(*
    Pneumatic actuator, single or double acting, ported from the legacy
    FB_MotionPneumaticActuator. Implements I_PneumaticActuator. The limit switch state, the
    insert and retract exclusion and the output timeout come from FB_PneumaticCore, which
    FB_MPA uses as well.

    Position state from the limit switches (in = inserted LS, out = retracted LS):
        in AND out         INVALID
        NOT in AND out     RETRACTED
        in AND NOT out     INSERTED
        NOT in AND NOT out MOVING
    bDone: the commanded direction has reached its limit switch. bBusy: a command
    is active and its limit switch is not reached. xMPS_OK is TRUE only when the
    state is RETRACTED or INSERTED. The fast fault (device 'MPA', type code
    E_MotionFFType.PNEUMATIC_MOVE) trips when xMPS_OK is FALSE.

    Insert and retract requests are mutually exclusive: both set at once clears both.
    Single acting: ibSingleCntrl TRUE and ibCntrlHold TRUE keeps the output on after
    arrival. Double acting: both FALSE, the output drops once the limit switch of the
    commanded direction has been active for LimitSwitchLatchDuration (default 1 s).
    An output that does not reach its limit switch within TimeoutDuration (default
    10 s) sets bError and sErrorMessage until bReset is set.

    Legacy behaviour kept as is: ibPMPS_OK and ibOverrideInterlock are unused (PMPS
    permission is not implemented), and LogEvents (legacy ACT_Logger) is never called by the body.
*)
FUNCTION_BLOCK FB_PneumaticActuator IMPLEMENTS I_PneumaticActuator
VAR_INPUT
    // Actuator can be inserted
    ibInsertOK : BOOL;
    // Actuator can be retracted
    ibRetractOK : BOOL;
    // To be linked to the arbiter bit (unused, as in the legacy FB)
    ibPMPS_OK : BOOL;
    // TRUE if the actuator needs one output (single acting), FALSE if it needs two
    ibSingleCntrl : BOOL;
    // Output must keep its value. TRUE for single acting, FALSE for double acting
    ibCntrlHold : BOOL;
    // If TRUE interlocks are ignored (unused, as in the legacy FB)
    ibOverrideInterlock : BOOL;
    {attribute 'pytmc' := '
    pv: FFO_Reset
    '}
    i_xReset : BOOL;
    {attribute 'pytmc' := '
    pv: FFO_AutoReset
    '}
    i_xAutoReset : BOOL;
END_VAR
VAR_OUTPUT
    {attribute 'pytmc' := '
    pv:
    '}
    stPneumaticActuator : ST_PneumaticActuator;
    {attribute 'pytmc' := '
     pv: MPS_OK
     field: ZNAM FALSE
     field: ONAM TRUE
     field: DESC TRUE if MPS signal is OK
    '}
    xMPS_OK : BOOL;
END_VAR
VAR
    // Fast fault output the fault is raised on
    fbFFHWO : REFERENCE TO FB_HardwareFFOutput;
    // Fault occurs while the actuator is not at a limit switch
    fbFF : FB_FastFault := (
        i_DevName := 'MPA',
        i_Desc := 'Fault occurs when the device is moving',
        i_TypeCode := E_MotionFFType.PNEUMATIC_MOVE);

    ftInit : R_TRIG;
    bFirstPass : BOOL;

    // Shared behaviour of the pneumatic actuator blocks
    fbCore : FB_PneumaticCore;
    // Time an output may stay on without reaching its limit switch
    tTimeOutDuration : TIME := T#10S;
    // Time a limit switch must stay active before a double acting output drops
    tLimitSwitchLatchDuration : TIME := T#1S;
    tonInsertLimitSwitch : TON;
    tonRetractLimitSwitch : TON;

    fbLogger : FB_LogMessage := (eSubsystem := E_SubSystem.MOTION);
    ePrevState : E_PnuematicActuatorPositionState;
    ftAction : R_TRIG;

    i_xInsertedLS AT %I* : BOOL;
    i_xRetractedLS AT %I* : BOOL;
    q_xInsert_DO AT %Q* : BOOL;
    q_xRetract_DO AT %Q* : BOOL;
END_VAR

IF NOT __ISVALIDREF(fbFFHWO) THEN
    RETURN;
END_IF

ftInit(CLK := TRUE, Q => bFirstPass);
IF bFirstPass THEN
    stPneumaticActuator.eState := E_PnuematicActuatorPositionState.INVALID;
    stPneumaticActuator.bRetractCmd := FALSE;
    stPneumaticActuator.bInsertCmd := FALSE;
END_IF

UpdateIO();

// Position state from the limit switches
// The output bits are those of the previous scan, so the timeout is reported one scan late
fbCore(
    bInLimitSwitch := stPneumaticActuator.bInLimitSwitch,
    bOutLimitSwitch := stPneumaticActuator.bOutLimitSwitch,
    bInsertOutput := stPneumaticActuator.bInsertOutput,
    bRetractOutput := stPneumaticActuator.bRetractOutput,
    tTimeout := tTimeOutDuration,
    eState => stPneumaticActuator.eState);

stPneumaticActuator.bDone := (stPneumaticActuator.bRetractCmd AND stPneumaticActuator.eState = E_PnuematicActuatorPositionState.RETRACTED)
    OR (stPneumaticActuator.bInsertCmd AND stPneumaticActuator.eState = E_PnuematicActuatorPositionState.INSERTED);
stPneumaticActuator.bBusy := (stPneumaticActuator.bRetractCmd AND stPneumaticActuator.eState <> E_PnuematicActuatorPositionState.RETRACTED)
    OR (stPneumaticActuator.bInsertCmd AND stPneumaticActuator.eState <> E_PnuematicActuatorPositionState.INSERTED);

// MPS faults when the actuator is in motion
xMPS_OK := (stPneumaticActuator.eState = E_PnuematicActuatorPositionState.RETRACTED)
    OR (stPneumaticActuator.eState = E_PnuematicActuatorPositionState.INSERTED);

// PMPS permission: yet to be implemented

// Insert and retract requests cannot both be active
IF stPneumaticActuator.bInsertCmd AND stPneumaticActuator.bRetractCmd THEN
    stPneumaticActuator.bInsertCmd := FALSE;
    stPneumaticActuator.bRetractCmd := FALSE;
END_IF

// Redundant: clear the opposite output and request when one output is active
IF stPneumaticActuator.bInsertOutput THEN
    stPneumaticActuator.bRetractOutput := FALSE;
    stPneumaticActuator.bRetractCmd := FALSE;
END_IF
IF stPneumaticActuator.bRetractOutput THEN
    stPneumaticActuator.bInsertOutput := FALSE;
    stPneumaticActuator.bInsertCmd := FALSE;
END_IF

stPneumaticActuator.bRetractOutput := stPneumaticActuator.bRetractOK
    AND stPneumaticActuator.bRetractCmd
    AND NOT stPneumaticActuator.bInsertCmd;
stPneumaticActuator.bInsertOutput := stPneumaticActuator.bInsertOK
    AND stPneumaticActuator.bInsertCmd
    AND NOT stPneumaticActuator.bRetractCmd;

// Double acting: drop the output once the actuator is seated in its limit switch
IF NOT ibSingleCntrl AND NOT ibCntrlHold THEN
    IF stPneumaticActuator.bRetractCmd
        AND stPneumaticActuator.bOutLimitSwitch
        AND tonRetractLimitSwitch.Q THEN
        stPneumaticActuator.bRetractOutput := FALSE;
    END_IF
    IF stPneumaticActuator.bInsertCmd
        AND stPneumaticActuator.bInLimitSwitch
        AND tonInsertLimitSwitch.Q THEN
        stPneumaticActuator.bInsertOutput := FALSE;
    END_IF
END_IF

tonInsertLimitSwitch(IN := stPneumaticActuator.bInLimitSwitch, PT := tLimitSwitchLatchDuration);
tonRetractLimitSwitch(IN := stPneumaticActuator.bOutLimitSwitch, PT := tLimitSwitchLatchDuration);

// Moving position timeout
IF fbCore.bInsertTimedOut THEN
    stPneumaticActuator.bError := TRUE;
    stPneumaticActuator.sErrorMessage := 'Actuator insert timeout';
ELSIF fbCore.bRetractTimedOut THEN
    stPneumaticActuator.bError := TRUE;
    stPneumaticActuator.sErrorMessage := 'Actuator retract timeout';
END_IF
stPneumaticActuator.bError R= stPneumaticActuator.bReset;

fbFF(
    i_xOK := xMPS_OK,
    i_xReset := i_xReset,
    i_xAutoReset := i_xAutoReset,
    io_fbFFHWO := fbFFHWO
);

UpdateIO();

PROPERTY Busy : BOOL
GET
Busy := stPneumaticActuator.bBusy;
END_GET
END_PROPERTY

(* Rebinds the fast fault output. Call from the CallAfterInit of an enclosing FB. *)
METHOD CallAfterInitActuator
VAR_INPUT
    fbFFHWO : REFERENCE TO FB_HardwareFFOutput;
END_VAR
THIS^.fbFFHWO REF= fbFFHWO;
END_METHOD

PROPERTY Done : BOOL
GET
Done := stPneumaticActuator.bDone;
END_GET
END_PROPERTY

PROPERTY Error : BOOL
GET
Error := stPneumaticActuator.bError;
END_GET
END_PROPERTY

// Text of the active timeout error
PROPERTY ErrorMessage : STRING
GET
ErrorMessage := stPneumaticActuator.sErrorMessage;
END_GET
END_PROPERTY

// Error reset request, the same bit as the reset PV
PROPERTY ErrorReset : BOOL
GET
ErrorReset := stPneumaticActuator.bReset;
END_GET
SET
stPneumaticActuator.bReset := ErrorReset;
END_SET
END_PROPERTY

(* Stores the mandatory fast fault output at instantiation. *)
METHOD FB_Init : BOOL
VAR_INPUT
    // TRUE: the retain variables are initialized (reset warm / reset cold)
    bInitRetains : BOOL;
    // TRUE: the instance will be copied to the copy code afterward (online change)
    bInCopyCode : BOOL;
    fbFFHWO : REFERENCE TO FB_HardwareFFOutput;
END_VAR
THIS^.fbFFHWO REF= fbFFHWO;
END_METHOD

METHOD Insert
VAR_INPUT
END_VAR
stPneumaticActuator.bInsertCmd := TRUE;
END_METHOD

// Insert request, the same bit Insert() raises. Write FALSE to clear it
PROPERTY InsertCmd : BOOL
GET
InsertCmd := stPneumaticActuator.bInsertCmd;
END_GET
SET
stPneumaticActuator.bInsertCmd := InsertCmd;
END_SET
END_PROPERTY

// Inserted limit switch input. Settable so tests and simulation can drive it
PROPERTY InsertedLS : BOOL
GET
InsertedLS := i_xInsertedLS;
END_GET
SET
i_xInsertedLS := InsertedLS;
END_SET
END_PROPERTY

// Insert digital output
PROPERTY InsertOutput : BOOL
GET
InsertOutput := q_xInsert_DO;
END_GET
END_PROPERTY

// Time a limit switch must stay active before a double acting output drops. Default 1 s
PROPERTY LimitSwitchLatchDuration : TIME
GET
LimitSwitchLatchDuration := tLimitSwitchLatchDuration;
END_GET
SET
tLimitSwitchLatchDuration := LimitSwitchLatchDuration;
END_SET
END_PROPERTY

(* Logs timeouts, insert and retract commands and state changes. Kept as in the
   legacy FB: the body does not call it. *)
METHOD LogEvents
// Log timeouts
IF fbCore.InsertTimeoutElapsed OR fbCore.RetractTimeoutElapsed THEN
    fbLogger(
        sMsg := stPneumaticActuator.sErrorMessage,
        eSevr := TcEventSeverity.Warning);
END_IF

// Log actuator commands
ftAction(CLK := stPneumaticActuator.bRetractOutput OR stPneumaticActuator.bInsertOutput);
IF ftAction.Q THEN
    IF stPneumaticActuator.bRetractOutput THEN
        fbLogger(
            sMsg := 'Actuator commanded retract',
            eSevr := TcEventSeverity.Info);
    END_IF
    IF stPneumaticActuator.bInsertOutput THEN
        fbLogger(
            sMsg := 'Actuator commanded insert',
            eSevr := TcEventSeverity.Info);
    END_IF
END_IF

// Log state changes
IF ePrevState <> stPneumaticActuator.eState THEN
    CASE stPneumaticActuator.eState OF
        E_PnuematicActuatorPositionState.INVALID:
            fbLogger(
                sMsg := 'Actuator invalid position.',
                eSevr := TcEventSeverity.Critical);
        E_PnuematicActuatorPositionState.MOVING:
            fbLogger(
                sMsg := 'Actuator moving',
                eSevr := TcEventSeverity.Warning);
        E_PnuematicActuatorPositionState.RETRACTED:
            fbLogger(
                sMsg := 'Actuator Retracted.',
                eSevr := TcEventSeverity.Info);
        E_PnuematicActuatorPositionState.INSERTED:
            fbLogger(
                sMsg := 'Actuator Inserted.',
                eSevr := TcEventSeverity.Info);
    END_CASE
    ePrevState := stPneumaticActuator.eState;
END_IF
END_METHOD

PROPERTY MpsOk : BOOL
GET
MpsOk := xMPS_OK;
END_GET
END_PROPERTY

METHOD Retract
VAR_INPUT
END_VAR
stPneumaticActuator.bRetractCmd := TRUE;
END_METHOD

// Retract request, the same bit Retract() raises. Write FALSE to clear it
PROPERTY RetractCmd : BOOL
GET
RetractCmd := stPneumaticActuator.bRetractCmd;
END_GET
SET
stPneumaticActuator.bRetractCmd := RetractCmd;
END_SET
END_PROPERTY

// Retracted limit switch input. Settable so tests and simulation can drive it
PROPERTY RetractedLS : BOOL
GET
RetractedLS := i_xRetractedLS;
END_GET
SET
i_xRetractedLS := RetractedLS;
END_SET
END_PROPERTY

// Retract digital output
PROPERTY RetractOutput : BOOL
GET
RetractOutput := q_xRetract_DO;
END_GET
END_PROPERTY

PROPERTY State : E_PnuematicActuatorPositionState
GET
State := stPneumaticActuator.eState;
END_GET
END_PROPERTY

// Time an output may stay on without reaching its limit switch. Default 10 s
PROPERTY TimeoutDuration : TIME
GET
TimeoutDuration := tTimeOutDuration;
END_GET
SET
tTimeOutDuration := TimeoutDuration;
END_SET
END_PROPERTY

(* Soft IO mapping: copies the limit switch inputs into the status struct, the
   command outputs into the digital outputs, and the interlock bits into the
   struct. Runs at the start and end of every body scan. *)
METHOD UpdateIO
// Inputs
stPneumaticActuator.bInLimitSwitch := i_xInsertedLS;
stPneumaticActuator.bOutLimitSwitch := i_xRetractedLS;

// Outputs
q_xInsert_DO := stPneumaticActuator.bInsertOutput;
q_xRetract_DO := stPneumaticActuator.bRetractOutput;

// EPICS
stPneumaticActuator.bRetractOK := ibRetractOK;
stPneumaticActuator.bInsertOK := ibInsertOK;
END_METHOD

END_FUNCTION_BLOCK

(* stored: Version 1.1.0.1
   POU FB_PneumaticActuator: Id {2f07bb5c-4a09-4cf3-874c-6ca5c05d35a8}, SpecialFunc None
   Property Busy: Id {9bc6d5a9-702c-47e7-8166-1ff1bf1a1058}
   Get Get: Id {558243f3-fc44-4d78-977b-d7c698f621b2}
   Method CallAfterInitActuator: Id {d4f39575-c492-4742-a42f-29167fd1a19f}
   Property Done: Id {53888b0c-796a-4245-8b1e-1dabf8118611}
   Get Get: Id {d2ff4d2e-d252-4f85-b4bd-65a712cbc7de}
   Property Error: Id {8404d4fe-ff22-4c3b-958c-f587f956d75f}
   Get Get: Id {a498d7b7-9e5e-4cf0-a2a9-9446879be052}
   Property ErrorMessage: Id {cc079e73-010e-4ac8-b70e-342f7c938ef6}
   Get Get: Id {8bd0509c-857d-4374-bd3f-a3d990f743ca}
   Property ErrorReset: Id {1fb44bda-b5e4-4db8-a6ae-d9d57053d2a6}
   Get Get: Id {1257d8fa-858a-40fc-9f3a-a03e969704b1}
   Set Set: Id {ff19a5e1-fc0c-448e-a1ac-69e10cd2a790}
   Method FB_Init: Id {dac1e0fe-6d03-496d-91c2-c314cf683124}
   Method Insert: Id {a33cb450-2ea7-4a10-9312-12390589f06f}
   Property InsertCmd: Id {df39559b-4075-4827-a23c-96d0b4b660a0}
   Get Get: Id {6ec1283a-9887-49a2-bff1-0d60fdd85b71}
   Set Set: Id {5c6cbdd8-67ed-4261-853f-dcd6e7a6f5c1}
   Property InsertedLS: Id {d50b4eb3-ae12-4eca-9f67-e090df9f3108}
   Get Get: Id {ea485854-f877-4192-ab40-5a385f18d333}
   Set Set: Id {5247fb4e-0dbd-4913-9100-258129e88869}
   Property InsertOutput: Id {ce818098-9e63-48fe-ad1e-4b0e10280a30}
   Get Get: Id {8c941bba-a2eb-4c74-80f5-d00d9a85b317}
   Property LimitSwitchLatchDuration: Id {15253413-d704-404d-8a3c-d865fc8362d2}
   Get Get: Id {eb7e98dc-a4e2-43de-bbb8-e9fdbc838711}
   Set Set: Id {1c1a16fc-46f8-4b5a-8046-8ea23c898e3b}
   Method LogEvents: Id {13872233-2ed3-4b1f-aa46-893d344f713d}
   Property MpsOk: Id {f1e56251-3052-4465-a343-5e527db84d31}
   Get Get: Id {834fba7d-bc63-4096-8553-84a44455d44b}
   Method Retract: Id {c6502e4a-23e6-4bc8-bdad-76fb44e83e7c}
   Property RetractCmd: Id {affaf238-45d1-4fcd-a1e6-f07f70369464}
   Get Get: Id {99d24730-1d7b-4978-8d16-ff3c3e3a65de}
   Set Set: Id {bc1d3d75-474a-40ae-ae93-e05d7402cf84}
   Property RetractedLS: Id {9bfc5da6-1e31-4e16-b573-11cb52db9b36}
   Get Get: Id {84a292e3-3f2d-4a68-b4a0-0e5923f21879}
   Set Set: Id {00eabfeb-cd40-49b6-a01f-8f06716f48ce}
   Property RetractOutput: Id {42776977-6a41-4fac-81de-856b16eab600}
   Get Get: Id {f7e3f2fc-6773-42ca-b59b-cd9cd4fe132a}
   Property State: Id {796b8ae2-ff6f-4a82-98d3-f17470befb7d}
   Get Get: Id {b50988d7-db5a-4efe-afeb-c177ea018b3b}
   Property TimeoutDuration: Id {583d0873-ceb5-41d1-a4c4-b8ed03dc4dc0}
   Get Get: Id {561597dc-1058-4d8e-a121-bc170eab9e4f}
   Set Set: Id {5ba17003-76d0-481a-89f5-5fae3cf1147b}
   Method UpdateIO: Id {60848ba4-a65f-4284-9cf1-48a0ecc8af78} *)
